Staubli VAL3: Algorithm4.dtx

public num nInverseMatrix1[4 4]
  [0,0] = 4.865664
  [0,1] = 0.229739
  [0,2] = 18.957284
  [1,0] = -2.180441
  [1,1] = 5.500387
  [1,2] = 4.336984
  [2,0] = -0.506536
  [2,1] = -1.473409
  [2,2] = -0.0709054
  [3,3] = 1
public num nMatrix1[4 4]
  [0,0] = 0.042143
  [0,1] = -0.196069
  [0,2] = -0.725376
  [1,0] = -0.0165157
  [1,1] = 0.0650218
  [1,2] = -0.43854
  [2,0] = 0.0421337
  [2,1] = 0.0495361
  [2,2] = 0.191493
  [3,3] = 1
public num nMatrix2[4 4]
  [0,0] = 1
  [1,1] = 1
  [2,2] = 1
  [3,0] = 6.816645
  [3,1] = 1120.929616
  [3,2] = 833.829369
  [3,3] = 1
public num nMatrix3[4 4]
  [0,0] = 4.865664
  [0,1] = 0.229739
  [0,2] = 18.957284
  [1,0] = -2.180441
  [1,1] = 5.500387
  [1,2] = 4.336984
  [2,0] = -0.506536
  [2,1] = -1.473409
  [2,2] = -0.0709054
  [3,0] = -2833.317475
  [3,1] = 4938.541162
  [3,2] = 4931.555835
  [3,3] = 1
public num nTeach_3_1[4 4]
  [0,0] = -0.702285
  [0,1] = -0.0819432
  [0,2] = -0.707164
  [1,0] = -0.115862
  [1,1] = 0.993265
  [1,2] = -3.24847E-05
  [2,0] = 0.702404
  [2,1] = 0.0819108
  [2,2] = -0.70705
  [3,0] = 1004.56
  [3,1] = -0.844997
  [3,2] = 227.853426
  [3,3] = 1
public num nTeach_3_2[4 4]
  [0,0] = -0.744428
  [0,1] = 0.279367
  [0,2] = -0.606449
  [1,0] = -0.0993466
  [1,1] = 0.85181
  [1,2] = 0.514345
  [2,0] = 0.66027
  [2,1] = 0.443142
  [2,2] = -0.606357
  [3,0] = 1011.376645
  [3,1] = -59.246821
  [3,2] = 211.566344
  [3,3] = 1
public num nTeach_3_3[4 4]
  [0,0] = -0.879562
  [0,1] = 0.475436
  [0,2] = 0.0182124
  [1,0] = 0.434368
  [1,1] = 0.786788
  [1,2] = 0.438508
  [2,0] = 0.194153
  [2,1] = 0.393606
  [2,2] = -0.898543
  [3,0] = 1061.682795
  [3,1] = -69.818944
  [3,2] = 189.439756
  [3,3] = 1
frame fFrame = {fatherId=world[0]}
num nTeach_2_1[4 4]
num nTeach_2_2[4 4]
